(*
	Batch processor. onEmit enriches and stores records only. Call the FB body
	cyclically to advance the exporter and export the oldest queued records when
	the schedule delay elapses or a full batch is available.
*)
FUNCTION_BLOCK FB_LogRecordProcessor_Batch EXTENDS FB_LogRecordProcessor_Base;
VAR_OUTPUT
	scheduledDelayMillis: UDINT := 1000;	// maximum delay before queued records are exported
	maxExportBatchSize: UDINT := 512;		// maximum records transferred to one export
	lastOperationSucceeded: BOOL := TRUE;
	failureResult: E_LogRecordProcessorFailureReason;
END_VAR
VAR
	_scheduleDelayTimer: TON;
	_records: FB_LogRecordQueue(maxCount:=0);  // set again during THIS^.FB_Init
	_exporter: REFERENCE TO FB_LogRecordExporter_Base;
	_rejectedCount: UDINT;  // records that could not be cloned or queued
END_VAR

// no-op; override to change log mutation/enrichment functionality
METHOD enrich
VAR_IN_OUT
	logRecord: FB_LogRecord;
END_VAR
END_METHOD

METHOD exportIfNeeded
VAR
	_exportFailureReason: E_LogRecordExporterFailureReason;
END_VAR
IF THIS^.maxExportBatchSize = 0
	OR_ELSE NOT __ISVALIDREF(THIS^._exporter)
	OR_ELSE THIS^._exporter.isBusy()
	OR_ELSE THIS^._records.count = 0 THEN
	RETURN;
END_IF

IF NOT THIS^._scheduleDelayTimer.Q
	AND_THEN THIS^._records.count < THIS^.maxExportBatchSize THEN
	RETURN;
END_IF

IF THIS^._exporter.export(
	logRecords:=THIS^._records,
	count:=THIS^.maxExportBatchSize,
	failureReason=>_exportFailureReason
) THEN
	THIS^._scheduleDelayTimer(IN:=FALSE, PT:=UDINT_TO_TIME(THIS^.scheduledDelayMillis));
	THIS^.lastOperationSucceeded := TRUE;
	THIS^.failureResult := E_LogRecordProcessorFailureReason.NA;
ELSE
	THIS^.lastOperationSucceeded := FALSE;
	THIS^.failureResult := E_LogRecordProcessorFailureReason.EXPORT_FAILURE;
END_IF
END_METHOD

METHOD FB_Exit : BOOL
VAR_INPUT
	bInCopyCode: BOOL;
END_VAR
IF NOT bInCopyCode THEN
	THIS^.free();
END_IF
END_METHOD

//FB_Init is always available implicitly and it is used primarily for initialization.
//The return value is not evaluated. For a specific influence, you can also declare the
//methods explicitly and provide additional code there with the standard initialization
//code. You can evaluate the return value.
METHOD FB_Init: BOOL
VAR_INPUT
    bInitRetains: BOOL; // TRUE: the retain variables are initialized (reset warm / reset cold)
    bInCopyCode: BOOL;  // TRUE: the instance will be copied to the copy code afterward (online change)
	maxQueueSize: UDINT := 2048;			// zero is unbounded; otherwise the oldest record is dropped when full
	scheduledDelayMillis: UDINT := 1000;	// maximum delay before queued records are exported
	maxExportBatchSize: UDINT := 512;		// maximum records transferred to one export
	exporter: REFERENCE TO FB_LogRecordExporter_Base;	// the exporter where the LogRecords are pushed.
END_VAR
THIS^._records.FB_Init(FALSE, FALSE, maxQueueSize);
THIS^.scheduledDelayMillis := scheduledDelayMillis;
THIS^.maxExportBatchSize := maxExportBatchSize;
IF __ISVALIDREF(exporter) THEN
	THIS^._exporter REF= exporter;
END_IF
END_METHOD

METHOD free
THIS^._records.free();
THIS^._scheduleDelayTimer(IN:=FALSE, PT:=UDINT_TO_TIME(THIS^.scheduledDelayMillis));
END_METHOD

(*
	Clones the log record onto the tail of the arrival-order queue.
	When the queue holds maxQueueSize records, the oldest record is
	dropped from the head to make room for the newest.
*)
METHOD onEmit
VAR_INPUT
	logRecord: REFERENCE TO FB_LogRecord;
END_VAR
VAR
	_pRecord: POINTER TO FB_LogRecord;
	_cloneFailureResult: E_LogRecordCloneFailureReason;
	_queueFailureReason: E_LogRecordQueueFailureReason;
END_VAR
THIS^.enrich(logRecord);

IF __ISVALIDREF(THIS^._exporter) THEN
	_pRecord := 0;
	IF NOT logRecord.cloneTo(pDest:=_pRecord, failureReason=>_cloneFailureResult) THEN
		IF _pRecord <> 0 THEN _pRecord^.delete(pSelf:=_pRecord); END_IF
		THIS^._rejectedCount := THIS^._rejectedCount + 1;
		THIS^.lastOperationSucceeded := FALSE;
		THIS^.failureResult := E_LogRecordProcessorFailureReason.RECORD_CLONE_FAILURE;
		RETURN;
	END_IF
	
	IF NOT THIS^._records.push(pValue:=_pRecord, failureReason=>_queueFailureReason) THEN
		_pRecord^.delete(pSelf:=_pRecord);
		THIS^._rejectedCount := THIS^._rejectedCount + 1;
		THIS^.lastOperationSucceeded := FALSE;
		THIS^.failureResult := E_LogRecordProcessorFailureReason.QUEUE_PUSH_FAILURE;
		RETURN;
	END_IF
END_IF

THIS^.lastOperationSucceeded := TRUE;
THIS^.failureResult := E_LogRecordProcessorFailureReason.NA;
END_METHOD

METHOD tick
VAR
	_exportFailureReason: E_LogRecordExporterFailureReason;
END_VAR
THIS^._scheduleDelayTimer(
	IN:=THIS^._records.count > 0,
	PT:=UDINT_TO_TIME(THIS^.scheduledDelayMillis)
);

IF __ISVALIDREF(THIS^._exporter) THEN
	THIS^._exporter.tick(failureReason=>_exportFailureReason);
	THIS^.exportIfNeeded();
END_IF
END_METHOD

(* Records lost so far: evicted from a full queue, or not cloned or queued. *)
PROPERTY droppedCount : UDINT
GET
droppedCount := THIS^._records.droppedCount + THIS^._rejectedCount;
END_GET
END_PROPERTY

(* Records waiting for export. *)
PROPERTY queuedCount : UDINT
GET
queuedCount := THIS^._records.count;
END_GET
END_PROPERTY

END_FUNCTION_BLOCK

(* stored: Version 1.1.0.1
   POU FB_LogRecordProcessor_Batch: Id {3c63b4ac-33ba-4480-a899-f0c3be47a7cf}, SpecialFunc None
   Method enrich: Id {cd91d31c-cfa3-4b93-ac03-7d361155ee3a}
   Method exportIfNeeded: Id {12d3e85a-6355-4c3e-8fcb-622a0ed4c3c0}
   Method FB_Exit: Id {ee6e60b0-3b81-40b7-905a-5fd33600daae}
   Method FB_Init: Id {1b6c3aba-d3d8-44a7-8d93-ac13d7ad0810}
   Method free: Id {f13c14df-6aac-4e5f-ae77-f40c30ac792c}
   Method onEmit: Id {601f420a-eb68-4a65-8062-d11e0d96dc3c}
   Method tick: Id {52431084-38a6-4b97-9c40-41396451732f}
   Property droppedCount: Id {ed729752-7b74-4e0a-9963-6ad4aaec6062}
   Get Get: Id {47f1e96e-54ee-453d-a0d3-809aa8416382}
   Property queuedCount: Id {98393c3e-b6b5-44af-b991-f83094a1eeb9}
   Get Get: Id {d0c264ce-15f6-43dd-a92b-238b6beb096c} *)
